(* IEC 61131-3 sources: P26002_Bosch_HDPump/P26002_Bosch_HDPump_PLC/DeviceFBs, 6 files *)

(* ---- FB_CAN_Broker_Modular.st ---- *)
(********************************************************************************
 * FUNCTION_BLOCK: FB_CAN_Broker_Modular
 *
 * Beschreibung:
 *   Vollständig modularer Hardware-Treiber-Manager für den CAN-Bus an Bachmann M1.
 *
 *   Vorteile:
 *     1. Dynamische Kanalanzahl: Über den Input 'NumChannels' wird festgelegt,
 *        wie viele Kanäle (1..16) aktiv genutzt werden.
 *     2. Vorgegebene Konfigurationstabelle ("Maske"):
 *        Alle CAN-IDs werden in einem Array 'Channels' übergeben.
 *     3. Automatische Schleifenabarbeitung:
 *        - Schaltet alle konfigurierten RxCobIds automatisch beim CAN-Controller frei.
 *        - Verteilt eintreffende Telegramme dynamisch auf den passenden Kanal.
 *        - Faires Round-Robin Sende-Management über alle aktiven Kanäle.
 *     4. Universelle Telegrammlänge (Msg_Length >= 1):
 *        Auch kurze Frames (1 Byte oder 2 Bytes) werden zuverlässig verarbeitet.
 ********************************************************************************)
FUNCTION_BLOCK FB_CAN_Broker_Modular
VAR_INPUT
    Enable          : BOOL := TRUE;             (* Broker aktivieren *)
    Reset           : BOOL := FALSE;            (* Re-Init auslösen *)
    NetNb           : DINT := 1;                (* CAN NetNumber (Standard: 1) *)
    CardNb          : DINT := 2;                (* CPU Card Number (Card 2) *)
    Chan            : UDINT := 0;               (* CAN-Kanal (0 = CAN A) *)
    NumChannels     : INT := 5;                 (* Anzahl der aktiv genutzten Kanäle (1..32) *)
END_VAR

VAR_IN_OUT
    (* Konfigurationstabelle / Maske aller Kanäle *)
    Channels        : ARRAY [1..32] OF ST_CAN_Broker_Channel;
END_VAR

VAR_OUTPUT
    Ready           : BOOL := FALSE;            (* Treiber initialisiert & betriebsbereit *)
    Error           : BOOL := FALSE;            (* Hardware- oder Konfigurationsfehler *)
    ErrorID         : DINT := 0;
    ActiveCount     : INT := 0;                 (* Tatsächlich überwachte Kanäle *)
END_VAR

VAR
    initStep        : INT := 0;
    initDone        : BOOL := FALSE;

    (* CUL Instanzen *)
    fbAttachEvent   : CUL_AttachEvent;
    fbSendMsg       : CUL_SendMsg_NB;
    fbRecvMsg       : CUL_ReceiveMsg;

    dwEventFlags    : UDINT := 0;
    nRet            : DINT := 0;

    (* Dynamische Rx-ID-Registrierung *)
    lastEnabledRx   : ARRAY [1..32] OF UDINT;

    (* Sende-Verwaltung *)
    txActive        : BOOL := FALSE;
    activeChan      : INT := 0;
    lastServedChan  : INT := 1;
    currTxCobId     : UDINT := 0;
    currTxData      : ARRAY [0..7] OF BYTE;

    (* Hilfsvariablen *)
    i               : INT;
    nActive         : INT;
    candChan        : INT;
    rxCount         : INT;
END_VAR

(* Begrenzung der aktiven Kanalanzahl auf 1..32 *)
nActive := NumChannels;
IF nActive < 1 THEN
    nActive := 1;
ELSIF nActive > 32 THEN
    nActive := 32;
END_IF;
ActiveCount := nActive;

(* ============================================================================ *)
(* Deaktivierung & Reset                                                       *)
(* ============================================================================ *)
IF NOT Enable THEN
    IF initDone THEN
        Cul_DetachEvent(NetNb := NetNb, Event := 0);
    END_IF;
    Ready    := FALSE;
    initDone := FALSE;
    initStep := 0;
    txActive := FALSE;
    RETURN;
END_IF;

IF Reset THEN
    IF initDone THEN
        Cul_DetachEvent(NetNb := NetNb, Event := 0);
    END_IF;
    Ready          := FALSE;
    Error          := FALSE;
    ErrorID        := 0;
    initDone       := FALSE;
    initStep       := 0;
    txActive       := FALSE;
    FOR i := 1 TO 32 DO
        lastEnabledRx[i] := 0;
    END_FOR;
END_IF;

(* ============================================================================ *)
(* Initialisierung der Hardware (Schritt 0)                                     *)
(* ============================================================================ *)
IF NOT initDone THEN
    CASE initStep OF
        0:
            (* Alle aktiven RxCobIds beim CAN-Controller freischalten *)
            FOR i := 1 TO nActive DO
                IF Channels[i].RxCobId > 0 AND Channels[i].RxCobId <> lastEnabledRx[i] THEN
                    nRet := Cul_EnableMsg(CardNb := CardNb, Chan := Chan, CobId := Channels[i].RxCobId);
                    lastEnabledRx[i] := Channels[i].RxCobId;
                END_IF;
            END_FOR;

            dwEventFlags := 0;
            fbAttachEvent(Req := TRUE, NetNb := NetNb, Event := dwEventFlags);

            IF fbAttachEvent.Done THEN
                fbAttachEvent(Req := FALSE, NetNb := NetNb, Event := dwEventFlags);
                initDone := TRUE;
                Ready    := TRUE;
                Error    := FALSE;
                ErrorID  := 0;
            ELSIF fbAttachEvent.Error THEN
                Error    := TRUE;
                ErrorID  := fbAttachEvent.Status;
            END_IF;
    END_CASE;
    RETURN;
END_IF;

(* Nachträglich veränderte RxCobIds dynamisch nachregistrieren *)
FOR i := 1 TO nActive DO
    IF Channels[i].RxCobId > 0 AND Channels[i].RxCobId <> lastEnabledRx[i] THEN
        nRet := Cul_EnableMsg(CardNb := CardNb, Chan := Chan, CobId := Channels[i].RxCobId);
        lastEnabledRx[i] := Channels[i].RxCobId;
    END_IF;
END_FOR;

(* ============================================================================ *)
(* Zyklus-Start: Flanken und Trigger der aktiven Kanäle zurücksetzen            *)
(* ============================================================================ *)
FOR i := 1 TO nActive DO
    Channels[i].RxNew   := FALSE;
    Channels[i].TxDone  := FALSE;
    Channels[i].TxError := FALSE;
END_FOR;

(* ============================================================================ *)
(* 1. EMPFANG: Hardware-Queue leeren & an Kanäle 1..nActive verteilen           *)
(* ============================================================================ *)
rxCount := 0;
REPEAT
    fbRecvMsg(NetNb := NetNb);
    rxCount := rxCount + 1;

    IF fbRecvMsg.Status = 0 AND fbRecvMsg.Msg_Length >= 1 THEN
        FOR i := 1 TO nActive DO
            IF Channels[i].RxCobId = fbRecvMsg.CobId THEN
                Channels[i].RxNew  := TRUE;
                Channels[i].RxData := fbRecvMsg.Msg_Data;
                Channels[i].RxLen  := fbRecvMsg.Msg_Length;
                EXIT;
            END_IF;
        END_FOR;
    END_IF;
UNTIL (fbRecvMsg.Status <> 0) OR (fbRecvMsg.Msg_Left = 0) OR (rxCount > 30)
END_REPEAT;

(* ============================================================================ *)
(* 2. SENDEN: Laufende Übertragung überwachen oder neuen Auftrag starten        *)
(* ============================================================================ *)
IF txActive THEN
    fbSendMsg(
        Req        := TRUE,
        NetNb      := NetNb,
        CobId      := currTxCobId,
        Msg_Data   := currTxData,
        Msg_Length := 8
    );

    IF fbSendMsg.Done THEN
        fbSendMsg(Req := FALSE, NetNb := NetNb, CobId := currTxCobId, Msg_Data := currTxData, Msg_Length := 8);
        txActive := FALSE;
        IF activeChan >= 1 AND activeChan <= nActive THEN
            Channels[activeChan].TxDone := TRUE;
            Channels[activeChan].TxBusy := FALSE;
            Channels[activeChan].TxReq  := FALSE;
        END_IF;
    ELSIF fbSendMsg.Error THEN
        fbSendMsg(Req := FALSE, NetNb := NetNb, CobId := currTxCobId, Msg_Data := currTxData, Msg_Length := 8);
        txActive := FALSE;
        IF activeChan >= 1 AND activeChan <= nActive THEN
            Channels[activeChan].TxError := TRUE;
            Channels[activeChan].TxBusy  := FALSE;
            Channels[activeChan].TxReq   := FALSE;
        END_IF;
    END_IF;

ELSE
    (* Round-Robin über alle nActive Kanäle *)
    FOR i := 1 TO nActive DO
        candChan := ((lastServedChan - 1 + i) MOD nActive) + 1;

        IF Channels[candChan].TxReq THEN
            activeChan                := candChan;
            lastServedChan            := candChan;
            currTxCobId               := Channels[candChan].TxCobId;
            currTxData                := Channels[candChan].TxData;
            Channels[candChan].TxBusy := TRUE;
            txActive                  := TRUE;
            EXIT;
        END_IF;
    END_FOR;

    IF txActive THEN
        fbSendMsg(
            Req        := TRUE,
            NetNb      := NetNb,
            CobId      := currTxCobId,
            Msg_Data   := currTxData,
            Msg_Length := 8
        );
    END_IF;
END_IF;

END_FUNCTION_BLOCK

(* ---- FB_CAN_Signal.st ---- *)
(********************************************************************************
 * FUNCTION_BLOCK: FB_CAN_Signal
 *
 * Beschreibung:
 *   Universeller Signal-Baustein zur Extraktion (Lesen / Decodieren) und
 *   Einbettung (Schreiben / Encodieren) von CAN-Signalen in das 8-Byte
 *   Nutzdatenfeld (Data) einer CAN-Nachricht.
 *
 *   Kompatibel mit Bachmann M-PLC (SolutionCenter):
 *     - Verwendet standardkonforme IEC 61131-3 Typkonvertierungen (<SOURCE>_TO_<TARGET>)
 *       (keine Kurzschreibweisen wie TO_UDINT, TO_DINT etc.).
 *     - Bit-Operationen (SHL, SHR, AND, OR, NOT) auf DWORD.
 *     - Entwickelt für Little-Endian (Intel-Format, Bosch Motorsport / RaceCon).
 ********************************************************************************)
FUNCTION_BLOCK FB_CAN_Signal
VAR_INPUT
    CobId       : UDINT := 0;       (* CAN Identifier (z. B. 16#650) zur Zuordnung/Doku *)
    StartBit    : UINT  := 0;       (* Start-Bit im CAN-Frame (0..63, LSB bei Little Endian) *)
    BitLength   : UINT  := 16;      (* Länge des Signals in Bits (1..32) *)
    IsSigned    : BOOL  := FALSE;   (* FALSE: Unsigned, TRUE: Signed *)
    Factor      : REAL  := 1.0;     (* Skalierungsfaktor: PhysValue = Raw * Factor + Offset *)
    Offset      : REAL  := 0.0;     (* Skalierungs-Offset *)
    bWrite      : BOOL  := FALSE;   (* FALSE = Lesen (Decode), TRUE = Schreiben (Encode) *)
    WriteValue  : REAL  := 0.0;     (* Zu schreibender physikalischer Wert (nur bei bWrite=TRUE) *)
END_VAR

VAR_IN_OUT
    Data        : ARRAY [0..7] OF BYTE; (* 8-Byte Nutzdatenfeld der CAN-Botschaft *)
END_VAR

VAR_OUTPUT
    RawValue    : UDINT := 0;       (* Extrahierter Rohwert als UDINT *)
    PhysValue   : REAL  := 0.0;     (* Skalierter physikalischer Messwert *)
    Valid       : BOOL  := FALSE;   (* Signal-Konfiguration gültig & Operation erfolgreich *)
    Error       : BOOL  := FALSE;   (* TRUE bei ungültigen Parametern (z.B. StartBit+Länge > 64) *)
END_VAR

VAR
    startByte   : UINT;
    bitOffset   : UINT;
    mask        : DWORD;
    signBit     : DWORD;
    dwRaw       : DWORD;
    dwRawWrite  : DWORD;
    nSignedVal  : DINT;
    rRawCalc    : REAL;
    i           : UINT;
    b           : UINT;
    currBitPos  : UINT;
    targetByte  : UINT;
    targetBit   : UINT;
    bitVal      : BOOL;
END_VAR

(* ============================================================================ *)
(* 1. Plausibilitätsprüfung der Signal-Parameter                                *)
(* ============================================================================ *)
IF (BitLength = 0) OR (BitLength > 32) OR ((StartBit + BitLength) > 64) THEN
    Error := TRUE;
    Valid := FALSE;
    RETURN;
END_IF;

Error := FALSE;
Valid := TRUE;

startByte := StartBit / 8;
bitOffset := StartBit MOD 8;

(* 32-Bit Bitmaske berechnen *)
IF BitLength >= 32 THEN
    mask := 16#FFFFFFFF;
ELSE
    mask := SHR(DWORD#16#FFFFFFFF, 32 - BitLength);
END_IF;

(* ============================================================================ *)
(* 2. SCHREIBEN (ENCODE): Signal in Data-Array einbetten                         *)
(* ============================================================================ *)
IF bWrite THEN
    IF Factor <> 0.0 THEN
        rRawCalc := (WriteValue - Offset) / Factor;
    ELSE
        rRawCalc := WriteValue;
    END_IF;

    nSignedVal := REAL_TO_DINT(rRawCalc);
    dwRawWrite := DINT_TO_DWORD(nSignedVal) AND mask;

    RawValue  := DWORD_TO_UDINT(dwRawWrite);
    PhysValue := WriteValue;

    (* Schnellpfad für byte-ausgerichtete Signale *)
    IF (bitOffset = 0) AND (BitLength = 8) THEN
        Data[startByte] := DWORD_TO_BYTE(dwRawWrite AND 16#FF);

    ELSIF (bitOffset = 0) AND (BitLength = 16) THEN
        Data[startByte]     := DWORD_TO_BYTE(dwRawWrite AND 16#FF);
        Data[startByte + 1] := DWORD_TO_BYTE(SHR(dwRawWrite, 8) AND 16#FF);

    ELSIF (bitOffset = 0) AND (BitLength = 24) THEN
        Data[startByte]     := DWORD_TO_BYTE(dwRawWrite AND 16#FF);
        Data[startByte + 1] := DWORD_TO_BYTE(SHR(dwRawWrite, 8) AND 16#FF);
        Data[startByte + 2] := DWORD_TO_BYTE(SHR(dwRawWrite, 16) AND 16#FF);

    ELSIF (bitOffset = 0) AND (BitLength = 32) THEN
        Data[startByte]     := DWORD_TO_BYTE(dwRawWrite AND 16#FF);
        Data[startByte + 1] := DWORD_TO_BYTE(SHR(dwRawWrite, 8) AND 16#FF);
        Data[startByte + 2] := DWORD_TO_BYTE(SHR(dwRawWrite, 16) AND 16#FF);
        Data[startByte + 3] := DWORD_TO_BYTE(SHR(dwRawWrite, 24) AND 16#FF);

    ELSE
        (* Universeller Pfad: Bitgenaues Read-Modify-Write *)
        FOR b := 0 TO (BitLength - 1) DO
            currBitPos := StartBit + b;
            targetByte := currBitPos / 8;
            targetBit  := currBitPos MOD 8;
            bitVal     := (SHR(dwRawWrite, b) AND 16#1) <> 16#0;

            IF targetByte <= 7 THEN
                IF bitVal THEN
                    Data[targetByte] := Data[targetByte] OR DWORD_TO_BYTE(SHL(DWORD#16#1, targetBit));
                ELSE
                    Data[targetByte] := Data[targetByte] AND NOT DWORD_TO_BYTE(SHL(DWORD#16#1, targetBit));
                END_IF;
            END_IF;
        END_FOR;
    END_IF;

    RETURN;
END_IF;

(* ============================================================================ *)
(* 3. LESEN (DECODE): Signal aus Data-Array extrahieren (Little Endian)        *)
(* ============================================================================ *)
(* Schnellpfad für byte-ausgerichtete Signale *)
IF (bitOffset = 0) AND (BitLength = 8) THEN
    dwRaw := BYTE_TO_DWORD(Data[startByte]);

ELSIF (bitOffset = 0) AND (BitLength = 16) THEN
    dwRaw := BYTE_TO_DWORD(Data[startByte]) OR SHL(BYTE_TO_DWORD(Data[startByte + 1]), 8);

ELSIF (bitOffset = 0) AND (BitLength = 24) THEN
    dwRaw := BYTE_TO_DWORD(Data[startByte])
          OR SHL(BYTE_TO_DWORD(Data[startByte + 1]), 8)
          OR SHL(BYTE_TO_DWORD(Data[startByte + 2]), 16);

ELSIF (bitOffset = 0) AND (BitLength = 32) THEN
    dwRaw := BYTE_TO_DWORD(Data[startByte])
          OR SHL(BYTE_TO_DWORD(Data[startByte + 1]), 8)
          OR SHL(BYTE_TO_DWORD(Data[startByte + 2]), 16)
          OR SHL(BYTE_TO_DWORD(Data[startByte + 3]), 24);

ELSE
    (* Universeller Pfad: Bis zu 5 Bytes zusammenführen und shiften *)
    dwRaw := 16#0;
    FOR i := 0 TO 3 DO
        IF (startByte + i) <= 7 THEN
            dwRaw := dwRaw OR SHL(BYTE_TO_DWORD(Data[startByte + i]), i * 8);
        END_IF;
    END_FOR;

    IF bitOffset > 0 THEN
        dwRaw := SHR(dwRaw, bitOffset);
        IF (startByte + 4) <= 7 THEN
            dwRaw := dwRaw OR SHL(BYTE_TO_DWORD(Data[startByte + 4]), 32 - bitOffset);
        END_IF;
    END_IF;

    dwRaw := dwRaw AND mask;
END_IF;

RawValue := DWORD_TO_UDINT(dwRaw);

(* ============================================================================ *)
(* 4. Vorzeichen-Erweiterung (Sign Extension) und Skalierung                    *)
(* ============================================================================ *)
IF IsSigned THEN
    signBit := SHL(DWORD#16#1, BitLength - 1);
    IF (dwRaw AND signBit) <> 16#0 THEN
        (* Negative Zahl: Führende Einsen auffüllen *)
        dwRaw := dwRaw OR (NOT mask);
    END_IF;
    nSignedVal := DWORD_TO_DINT(dwRaw);
    PhysValue  := (DINT_TO_REAL(nSignedVal) * Factor) + Offset;
ELSE
    nSignedVal := DWORD_TO_DINT(dwRaw);
    PhysValue  := (DINT_TO_REAL(nSignedVal) * Factor) + Offset;
END_IF;

END_FUNCTION_BLOCK

(* ---- FB_FuelSupply.st ---- *)
FUNCTION_BLOCK FB_FuelSupply
VAR_INPUT
HW_DI_FuelTank_Empty : BOOL;
SupplyFuelPumpPIDsettings: ARRAY [1..3] OF REAL;
SupplyFuelPump_pressure_tolerance : REAL;
END_VAR

VAR_OUTPUT
HW_DO_EnableAdjPowerSupply : BOOL;
HW_AO_FuelPumpSupplyVoltage : REAL;
END_VAR

VAR_IN_OUT
fbIO_FuelSupply : FuelSupply;
END_VAR

VAR
init : BOOL := FALSE;

max_fuelsupply_pressure : REAL := 10; (*bar*)

Enable : INT;
PID_Controller : Cont_PIDT1_Par;
TS : REAL := 1.0;
T1 : REAL := 0.0;
MaxOutput : REAL := 100.0;
MinOutput : REAL := 0.0;

END_VAR

fbIO_FuelSupply.pressure_tolerance := SupplyFuelPump_pressure_tolerance;
ACT_SET_PIDvalues;
IF NOT init THEN
	init := TRUE;
END_IF

(* ENABLE GATE *)

IF NOT fbIO_FuelSupply.enable THEN
	HW_DO_EnableAdjPowerSupply := FALSE;
	HW_AO_FuelPumpSupplyVoltage := 0.0;
	Enable := 0;
	RETURN;
ELSE
	Enable := 3;
END_IF

(* Pumpen anschalten *)
IF fbIO_FuelSupply.start THEN
	HW_DO_EnableAdjPowerSupply := TRUE;
	fbIO_FuelSupply.start := FALSE;
END_IF

(* Pumpen ausschalten *)
IF fbIO_FuelSupply.stop THEN
	HW_DO_EnableAdjPowerSupply := FALSE;
	fbIO_FuelSupply.stop := FALSE;
END_IF

fbIO_FuelSupply.running := HW_DO_EnableAdjPowerSupply;

(* Neuen Sollwert übernehmen *)

IF ABS(fbIO_FuelSupply.SV-fbIO_FuelSupply.SVreq) > 0.01 THEN

	IF fbIO_FuelSupply.SVreq < max_fuelsupply_pressure THEN
		fbIO_FuelSupply.SVaccepted := TRUE;
	ELSE
		fbIO_FuelSupply.SVaccepted := FALSE;
	END_IF

	IF fbIO_FuelSupply.SVaccepted THEN
		fbIO_FuelSupply.SV := fbIO_FuelSupply.SVreq;
	END_IF

END_IF

PID_Controller ( Enable := Enable, (* 0 - Regler deaktivieren;
 											  * 1 - Regler initialisieren (PValue, IValue, DValue und TS neu übernehmen);
 											  * 2 - Regler aktivieren;
 											  * 3 - Regler initialisieren und aktivieren (PValue, IValue, DValue und TS neu übernehmen und regeln)*)

                 SetValue := fbIO_FuelSupply.SV,
                 ActValue := fbIO_FuelSupply.AV,
                 PValue := fbIO_FuelSupply.PID[1],
                 IValue := fbIO_FuelSupply.PID[2],
                 DValue := fbIO_FuelSupply.PID[3],
                 TS := TS,
                 T1 := T1,
                 MaxOutput := MaxOutput,
                 MinOutput := MinOutput );

		fbIO_FuelSupply.pid_error     	:= PID_Controller.Error;
		HW_AO_FuelPumpSupplyVoltage    	:= PID_Controller.OutVar;

IF ABS(fbIO_FuelSupply.AV-fbIO_FuelSupply.SV) < fbIO_FuelSupply.pressure_tolerance THEN
	fbIO_FuelSupply.SVreached := TRUE;
ELSE
	fbIO_FuelSupply.SVreached := FALSE;
END_IF

;
END_FUNCTION_BLOCK

ACTIONS
	ACTION ACT_SET_PIDvalues
		IF fbIO_FuelSupply.setPID OR NOT init THEN
			fbIO_FuelSupply.PID[1] := SupplyFuelPumpPIDsettings[1];
			fbIO_FuelSupply.PID[2] := SupplyFuelPumpPIDsettings[2];
			fbIO_FuelSupply.PID[3] := SupplyFuelPumpPIDsettings[3];
			fbIO_FuelSupply.setPID := FALSE;
		END_IF
	END_ACTION

END_ACTIONS

(* ---- FB_MASS6000_DP.st ---- *)
(********************************************************************************
 * FUNCTION_BLOCK: FB_MASS6000_DP
 *
 * Beschreibung:
 *   Decodierung und Aufbereitung der PROFIBUS-DP / PROFINET Prozessdaten
 *   des Coriolis-Massendurchflussmessers Siemens SITRANS FC MASSFLO MASS 6000
 *   über das ADFweb PROFINET/PROFIBUS Gateway HD67604-A1.
 *
 *   Konfiguration: "Fall A" (4 Messwertmodule à 5 Byte = 20 Byte E/A)
 *   ----------------------------------------------------------------------------
 *   Offset (Bytes) | Messgröße          | Datentyp               | Umrechnung
 *   ----------------------------------------------------------------------------
 *   Byte 0..3      | Massflow (Masse)   | IEEE-754 Float (Big-E) | kg/s * 3600 -> kg/h
 *   Byte 4         | Status Massflow    | PA-Statusbyte (8 Bit)  | >= 16#80 = Good
 *   Byte 5..8      | Volumeflow (Vol.)  | IEEE-754 Float (Big-E) | m3/h bzw. l/h
 *   Byte 9         | Status Volumeflow  | PA-Statusbyte (8 Bit)  | >= 16#80 = Good
 *   Byte 10..13    | Density (Dichte)   | IEEE-754 Float (Big-E) | kg/l (1:1)
 *   Byte 14        | Status Density     | PA-Statusbyte (8 Bit)  | >= 16#80 = Good
 *   Byte 15..18    | Temperature (Temp) | IEEE-754 Float (Big-E) | Kelvin - 273.15 -> °C
 *   Byte 19        | Status Temperature | PA-Statusbyte (8 Bit)  | >= 16#80 = Good
 *
 *   Kompatibel mit Bachmann M-PLC (SolutionCenter):
 *     - Standardkonforme Konvertierungen (<SOURCE>_TO_<TARGET>).
 *     - Bit-rekonstruierte Float-Wandlung über ADR() und POINTER TO REAL.
 ********************************************************************************)
FUNCTION_BLOCK FB_MASS6000_DP
VAR_INPUT
    bEnable             : BOOL := TRUE;             (* Baustein-Aktivierung *)
    Data                : ARRAY [0..19] OF BYTE;    (* 20-Byte PROFINET Eingangsbereich *)
END_VAR

VAR_OUTPUT
    rMassflow_kgh       : REAL := 0.0;              (* Massendurchfluss [kg/h] *)
    rVolumeflow         : REAL := 0.0;              (* Volumendurchfluss [m3/h bzw. l/h] *)
    rDensity_kgl        : REAL := 0.0;              (* Dichte [kg/l] *)
    rTemperature_degC   : REAL := 0.0;              (* Kraftstofftemperatur [°C] *)

    (* PROFIBUS PA Qualitäts-Statusbytes (>= 16#80 = Good) *)
    byStatusMassflow    : BYTE := 16#00;
    byStatusVolumeflow  : BYTE := 16#00;
    byStatusDensity     : BYTE := 16#00;
    byStatusTemperature : BYTE := 16#00;

    bMassflowValid      : BOOL := FALSE;            (* Massflow-Status OK *)
    bVolumeflowValid    : BOOL := FALSE;            (* Volumeflow-Status OK *)
    bDensityValid       : BOOL := FALSE;            (* Density-Status OK *)
    bTemperatureValid   : BOOL := FALSE;            (* Temperature-Status OK *)
    bAllValid           : BOOL := FALSE;            (* Alle 4 Messwerte gültig *)
END_VAR

VAR
    dwRawFloat          : DWORD;
    pRealHelper         : POINTER TO REAL;
    rRawValue           : REAL;
END_VAR

IF NOT bEnable THEN
    rMassflow_kgh       := 0.0;
    rVolumeflow         := 0.0;
    rDensity_kgl        := 0.0;
    rTemperature_degC   := 0.0;
    bMassflowValid      := FALSE;
    bVolumeflowValid    := FALSE;
    bDensityValid       := FALSE;
    bTemperatureValid   := FALSE;
    bAllValid           := FALSE;
    RETURN;
END_IF;

pRealHelper := ADR(dwRawFloat);

(* ============================================================================ *)
(* 1. Massflow (Byte 0..3: IEEE-754 Big-Endian Float, Byte 4: Status)           *)
(* ============================================================================ *)
dwRawFloat := SHL(BYTE_TO_DWORD(Data[0]), 24) OR
              SHL(BYTE_TO_DWORD(Data[1]), 16) OR
              SHL(BYTE_TO_DWORD(Data[2]), 8)  OR
              BYTE_TO_DWORD(Data[3]);

rRawValue          := pRealHelper^;
rMassflow_kgh      := rRawValue * 3600.0; (* Umrechnung kg/s in kg/h *)
byStatusMassflow   := Data[4];
bMassflowValid     := (byStatusMassflow AND 16#C0) = 16#80; (* PA Quality Bit: Good *)

(* ============================================================================ *)
(* 2. Volumeflow (Byte 5..8: IEEE-754 Big-Endian Float, Byte 9: Status)         *)
(* ============================================================================ *)
dwRawFloat := SHL(BYTE_TO_DWORD(Data[5]), 24) OR
              SHL(BYTE_TO_DWORD(Data[6]), 16) OR
              SHL(BYTE_TO_DWORD(Data[7]), 8)  OR
              BYTE_TO_DWORD(Data[8]);

rVolumeflow        := pRealHelper^;
byStatusVolumeflow := Data[9];
bVolumeflowValid   := (byStatusVolumeflow AND 16#C0) = 16#80;

(* ============================================================================ *)
(* 3. Density (Byte 10..13: IEEE-754 Big-Endian Float, Byte 14: Status)         *)
(* ============================================================================ *)
dwRawFloat := SHL(BYTE_TO_DWORD(Data[10]), 24) OR
              SHL(BYTE_TO_DWORD(Data[11]), 16) OR
              SHL(BYTE_TO_DWORD(Data[12]), 8)  OR
              BYTE_TO_DWORD(Data[13]);

rDensity_kgl       := pRealHelper^; (* Direkt in kg/l *)
byStatusDensity    := Data[14];
bDensityValid      := (byStatusDensity AND 16#C0) = 16#80;

(* ============================================================================ *)
(* 4. Temperature (Byte 15..18: IEEE-754 Big-Endian Float, Byte 19: Status)     *)
(* ============================================================================ *)
dwRawFloat := SHL(BYTE_TO_DWORD(Data[15]), 24) OR
              SHL(BYTE_TO_DWORD(Data[16]), 16) OR
              SHL(BYTE_TO_DWORD(Data[17]), 8)  OR
              BYTE_TO_DWORD(Data[18]);

rRawValue           := pRealHelper^;
rTemperature_degC   := rRawValue - 273.15; (* Kelvin nach Celsius *)
byStatusTemperature := Data[19];
bTemperatureValid   := (byStatusTemperature AND 16#C0) = 16#80;

(* Gesamt-Gültigkeitsbit *)
bAllValid := bMassflowValid AND bVolumeflowValid AND bDensityValid AND bTemperatureValid;

END_FUNCTION_BLOCK

(* ---- FB_OilConditioning.st ---- *)
FUNCTION_BLOCK FB_OilConditioning
VAR_INPUT
HW_AI_OilTemperature : REAL;
HW_AI_OilPressure : REAL;
OilConditioning_pressure_tolerance : REAL;
OilConditioning_temperature_tolerance : REAL;
END_VAR

VAR_OUTPUT
HW_AO_OilPressure : REAL;
HW_DO_EnableOilFan: BOOL;
HW_DO_EnableOilConditioning: BOOL;
END_VAR

VAR_IN_OUT
fbIO_OilConditioning : OilConditioning;
END_VAR

VAR
max_oil_pressure : REAL := 10; (* bar *)
max_oil_temperature : REAL := 90; (* °C)*)
END_VAR

fbIO_OilConditioning.temperature_tolerance      := OilConditioning_temperature_tolerance;
fbIO_OilConditioning.pressure_tolerance         := OilConditioning_pressure_tolerance;

fbIO_OilConditioning.actualOil_pressure := HW_AI_OilPressure;
fbIO_OilConditioning.actualOil_temperature := HW_AI_OilTemperature;

(* ENABLE GATE *)

IF NOT fbIO_OilConditioning.enable THEN
	HW_DO_EnableOilConditioning := FALSE;
	HW_DO_EnableOilFan := FALSE;
	HW_AO_OilPressure := 0.0;
	fbIO_OilConditioning.pressure_SVaccepted := FALSE;
	fbIO_OilConditioning.temperature_SVaccepted := FALSE;
	RETURN;
END_IF

(* Pumpen anschalten *)
IF fbIO_OilConditioning.start THEN
	HW_DO_EnableOilConditioning := TRUE;
ELSE
	HW_DO_EnableOilConditioning := FALSE;
END_IF

(* Lüfter anschalten *)
IF (fbIO_OilConditioning.actualOil_temperature - fbIO_OilConditioning.setOil_temperature) > 3*fbIO_OilConditioning.temperature_tolerance
	OR fbIO_OilConditioning.actualOil_temperature > max_oil_temperature THEN
	HW_DO_EnableOilFan := TRUE;
ELSE
	HW_DO_EnableOilFan := FALSE;
END_IF

(* Neuen Sollwert übernehmen *)

IF ABS(fbIO_OilConditioning.setOil_pressure-HW_AO_OilPressure) > 0.01 THEN

	IF fbIO_OilConditioning.setOil_pressure < max_oil_pressure THEN
		fbIO_OilConditioning.pressure_SVaccepted := TRUE;
	ELSE
		fbIO_OilConditioning.pressure_SVaccepted := FALSE;
	END_IF

	IF fbIO_OilConditioning.pressure_SVaccepted THEN
		HW_AO_OilPressure := fbIO_OilConditioning.setOil_pressure;
	END_IF

END_IF

IF fbIO_OilConditioning.setOil_temperature < max_oil_temperature THEN
	fbIO_OilConditioning.temperature_SVaccepted := TRUE;
ELSE
	fbIO_OilConditioning.temperature_SVaccepted := FALSE;
END_IF

IF ABS(fbIO_OilConditioning.actualOil_temperature-fbIO_OilConditioning.setOil_temperature) < fbIO_OilConditioning.temperature_tolerance THEN
	fbIO_OilConditioning.temperature_SVreached := TRUE;
ELSE
	fbIO_OilConditioning.temperature_SVreached := FALSE;
END_IF

IF ABS(fbIO_OilConditioning.actualOil_pressure-fbIO_OilConditioning.setOil_pressure) < fbIO_OilConditioning.pressure_tolerance THEN
	fbIO_OilConditioning.pressure_SVreached := TRUE;
ELSE
	fbIO_OilConditioning.pressure_SVreached := FALSE;
END_IF

;
END_FUNCTION_BLOCK

(* start:	BOOL; *)
(* stop:	BOOL; *)
(* enabled: BOOL; *)
(*  *)
(* setOil_temperature: REAL; *)
(* setOil_pressure: REAL; *)
(*  *)
(* actualOil_temperature: REAL; *)
(* actualOil_pressure: REAL; *)
(*  *)
(* temperature_tolerance      : REAL := 2; *)
(* pressure_tolerance         : REAL := 0.5; *)
(*  *)
(* temperature_SVaccepted           : BOOL := FALSE; *)
(* temperature_SVreached            : BOOL := FALSE; *)
(*  *)
(* pressure_SVaccepted           : BOOL := FALSE; *)
(* pressure_SVreached            : BOOL := FALSE; *)

(* ---- FB_Thermostat.st ---- *)
FUNCTION_BLOCK FB_Thermostat
VAR_INPUT
SupplyFuelPump_temperature_tolerance : REAL;
END_VAR

VAR_OUTPUT

END_VAR

VAR_IN_OUT
fbIO_Thermostat : Thermostat;
END_VAR

VAR

END_VAR

(* Kommunikation aufbauen *)

(* Ist-Werte lesen *)
fbIO_Thermostat.SV_tolerance := SupplyFuelPump_temperature_tolerance;

(* Fehler auswerten *)

(* Neue Soll-Werte schreiben*)

(* enable               : BOOL := FALSE;           (* Freigabe der Ansteuerung *) *)
(* card_nb              : INT := 0;                (* Steckplatz (Slot) der RS232-Karte am Bachmann Rack *) *)
(* chan_nb              : INT := 1;                (* Kanalnummer der RS232-Schnittstelle (1 oder 2) *) *)
(* baud_rate            : DINT := 9600;            (* Baudrate (Huber Standard: 9600) *) *)
(* state                : state_device := DV_INIT; (* Aktueller Gerätestatus gemäß state_device.dt *) *)
(* reset                : BOOL := FALSE;           (* Trigger: Fehler quittieren & zurücksetzen *) *)
(* start                : BOOL := FALSE;           (* Temperierung/Umwälzung starten (Mode 'C') *) *)
(* stop                 : BOOL := FALSE;           (* Temperierung/Umwälzung stoppen (Mode 'O') *) *)
(* set_setpoint         : BOOL := FALSE;           (* Trigger: Neuen Sollwert an Thermostat senden *) *)
(* target_setpoint      : REAL := 20.0;            (* Sollwert-Vorgabe in °C (z.B. 25.5 °C) *) *)
(* act_setpoint         : REAL := 0.0;             (* Rückgelesener Sollwert vom Thermostat in °C *) *)
(* temp_internal        : REAL := 0.0;             (* Interner Istwert F1 in °C *) *)
(* temp_external        : REAL := 0.0;             (* Externer Istwert F2 in °C (-151.00 = nicht vorhanden) *) *)
(* sensor_ext_connected : BOOL := TRUE;            (* FALSE = Externer Fühler F2 nicht angeschlossen/defekt *) *)
(* control_active       : BOOL := FALSE;           (* TRUE = Temperierung/Umwälzung aktiv *) *)
(* SVaccepted           : BOOL := FALSE;           (* TRUE = Sollwert vom Thermostat übernommen *) *)
(* SVreached            : BOOL := FALSE;           (* TRUE = Sollwert innerhalb Toleranz erreicht *) *)
(* SV_tolerance         : REAL := 0.5;             (* Toleranzband in °C für SVreached *) *)
(* device_alarm         : BOOL := FALSE;           (* TRUE = Gerät meldet Alarmstatus ('1') *) *)
(* watchdog_error       : BOOL := FALSE;           (* TRUE = Watchdog Timeout aufgetreten *) *)
(* com_status           : STRING := 'disconnected'; *)
(* com_ready            : BOOL := FALSE; *)
(*		 *)
;
END_FUNCTION_BLOCK
